(* PLC project TBEN_L5_PLC11.project, CODESYS CODESYS V3.5 SP21 Patch 1 *)
(* stored: creationDateTime 2026-11-07T15:35:08.6454114, modificationDateTime 2026-11-07T15:09:07.4034196 *)

// Chuyển StringT IO-Link (không có ký tự kết thúc) thành STRING, cắt ở 64 ký tự
FUNCTION F_IolBytesToStr : STRING(64)
VAR_INPUT
    pBuf  : POINTER TO BYTE;
    uiLen : UINT;
END_VAR
VAR
    sTmp : STRING(64);
    pDst : POINTER TO BYTE;
    i    : UINT;
    n    : UINT;
END_VAR

            sTmp := '';
IF pBuf <> 0 THEN
    n := MIN(uiLen, 64);
    pDst := ADR(sTmp);
    i := 0;
    WHILE i < n DO
        IF pBuf[i] = 0 THEN          // device có thể đệm 0 ở cuối
            EXIT;
        END_IF
        pDst[i] := pBuf[i];
        i := i + 1;
    END_WHILE
    pDst[i] := 0;
END_IF
F_IolBytesToStr := sTmp;

          
END_FUNCTION
